Fanuc KAREL source: ka00142.KL

-- PROVISIONAL review KL for V770-1; original PC SHA256 9d7e340cf36b73797bd3752b6ead82da2213b34c8aebec33d7f9a86fcbaa222a
-- Incomplete behavior may be omitted. Consult companion uncertainty JSON. Do not deploy.
PROGRAM KA00142
%NOLOCKGROUP
-- UNRESOLVED_DECL SRC type=002017
-- UNRESOLVED_DECL DST type=00001c
BEGIN
  -- UNRESOLVED_PC offsets 5-19; opcodes 2E,22,9D,33,B4
  -- UNRESOLVED_PC offsets 24-39; opcodes 22,9D,33,B3,23
  -- UNRESOLVED_PC offsets 44-48; opcodes 7F
END KA00142
